FUNCTION_BLOCK EQ_Crimper (* An equipment block: the only block that touches this equipment's pins. Skills send it what to switch over a local channel; it switches the outputs (off first, then on), reads the inputs every cycle and reports them to the skills and to OPC UA. One skill holds it at a time; on release or when the module aborts it switches everything off. Technical: Crimping head that closes around the cap; simulated until it is chosen (no pin on the Pi yet); equipment IO: owns its IO points, writes the output values its holder sends, reads its inputs every cycle and reports changes *)
  (* Standard: 61499-2 *)
  (* Version 0.1, 2026-09-28, Project contributors, AAU Smart Production Lab *)
  PACKAGE capping;
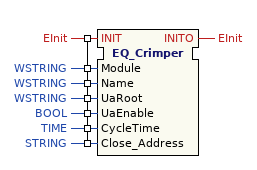
  EVENT_INPUT
    INIT : EInit WITH Module, Name, UaRoot, UaEnable, CycleTime, Close_Address; (* Initialise, once at start-up (the INIT chain); takes the values given with it *)
  END_EVENT
  EVENT_OUTPUT
    INITO : EInit; (* Initialised: the next block of the INIT chain goes on *)
  END_EVENT
  VAR_INPUT
    Module : WSTRING; (* The module's name; its local channels are named after it (loc[<Module>/...]) *)
    Name : WSTRING := "Crimper"; (* The equipment item's name: its local channels and OPC UA folder *)
    UaRoot : WSTRING; (* The module's OPC UA folder, e.g. /Objects/Filling *)
    UaEnable : BOOL; (* Publish on OPC UA *)
    CycleTime : TIME := T#50ms; (* How often the inputs are read *)
    Close_Address : STRING; (* Where Close is: 'gpio[chip:line(:pull_up|:pull_down)(:active_low)]', 'pwm[chip:channel:period_ns]', 'modbus[...]', 'sim', or an IO handle's name; empty: not connected *)
  END_VAR
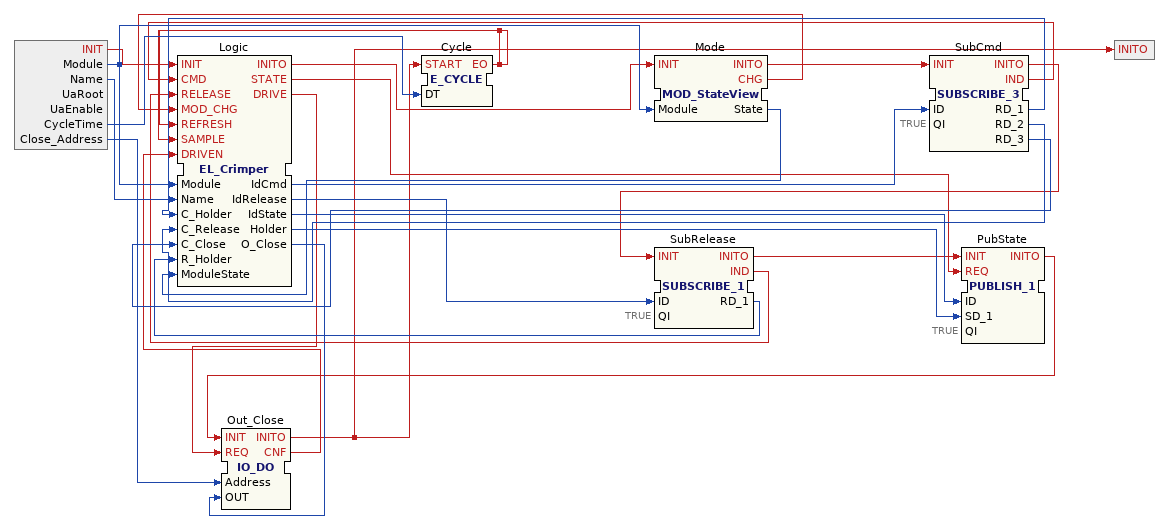
  (* Group Core: One holder at a time, break before make, all off on release or abort; scanned every CycleTime *)
  (* Group Channels: Local channels to and from the skills (cmd, release, state), the module's state, and the inputs over OPC UA *)
  (* Group Outputs: The equipment's actuators: written on a change and every cycle, one block per IO point *)
  FBS
    Logic : capping::EL_Crimper; (* The equipment's logic (EL_): takes commands from one holder at a time, switches the outputs (off first, then on), switches all off on release or module abort, and reports input changes. *) {SET_ATTRIBUTE(GroupName, Core)}
    Cycle : iec61499::events::E_CYCLE; (* Ticks every cycle so the inputs are read and the outputs refreshed. *) {SET_ATTRIBUTE(GroupName, Core)}
    Mode : modlib::MOD_StateView; (* Watches the module's PackML state, to switch everything off when the module aborts. *) {SET_ATTRIBUTE(GroupName, Channels)}
    SubCmd : iec61499::net::SUBSCRIBE_3(QI := TRUE); (* Receives the commands skills send on this equipment's command channel. *) {SET_ATTRIBUTE(GroupName, Channels)}
    SubRelease : iec61499::net::SUBSCRIBE_1(QI := TRUE); (* Hears the module's release channel: when its holder gives up, everything goes off. *) {SET_ATTRIBUTE(GroupName, Channels)}
    PubState : iec61499::net::PUBLISH_1(QI := TRUE); (* Publishes the inputs and the holder on this equipment's state channel, for the skills. *) {SET_ATTRIBUTE(GroupName, Channels)}
    Out_Close : modlib::IO_DO; (* The pin Close: switches the output at Close_Address (a Pi pin, Modbus, or simulated). *) {SET_ATTRIBUTE(GroupName, Outputs)}
  END_FBS
  EVENT_CONNECTIONS
    INIT TO Logic.INIT;
    Logic.INITO TO Mode.INIT;
    Mode.INITO TO SubCmd.INIT;
    SubCmd.INITO TO SubRelease.INIT;
    SubRelease.INITO TO PubState.INIT;
    PubState.INITO TO Out_Close.INIT;
    Out_Close.INITO TO Cycle.START;
    Out_Close.INITO TO INITO;
    SubCmd.IND TO Logic.CMD;
    SubRelease.IND TO Logic.RELEASE;
    Mode.CHG TO Logic.MOD_CHG;
    Cycle.EO TO Logic.REFRESH;
    Cycle.EO TO Logic.SAMPLE;
    Logic.STATE TO PubState.REQ;
    Logic.DRIVE TO Out_Close.REQ;
    Out_Close.CNF TO Logic.DRIVEN;
  END_CONNECTIONS
  DATA_CONNECTIONS
    Module TO Logic.Module;
    Name TO Logic.Name;
    Module TO Mode.Module;
    Logic.IdCmd TO SubCmd.ID;
    Logic.IdRelease TO SubRelease.ID;
    Logic.IdState TO PubState.ID;
    CycleTime TO Cycle.DT;
    SubCmd.RD_1 TO Logic.C_Holder;
    SubCmd.RD_2 TO Logic.C_Release;
    SubCmd.RD_3 TO Logic.C_Close;
    SubRelease.RD_1 TO Logic.R_Holder;
    Mode.State TO Logic.ModuleState;
    Logic.Holder TO PubState.SD_1;
    Close_Address TO Out_Close.Address;
    Logic.O_Close TO Out_Close.OUT;
  END_CONNECTIONS
END_FUNCTION_BLOCK
